(*
	Contract shared by span exporters. A processor offers a batch with export, which moves up to
	count of the oldest spans out of the processor's queue into the exporter without cloning
	them. The exporter owns the batch until free, which runs when the batch is delivered or
	failed, when the next batch is accepted, and when the exporter is destroyed.
	Concrete exporters advance delivery in tick and report through isBusy whether they can take
	another batch. Only ended spans reach an exporter.
*)
FUNCTION_BLOCK ABSTRACT FB_SpanExporter_Base
VAR
	_spans: FB_SpanQueue(maxCount:=0);
	_exportActive: BOOL;
	_callFailureReason: E_SpanExporterFailureReason;
END_VAR

(*
	Takes ownership of up to count of the oldest spans in spans. While busy it refuses with
	ACTIVE_EXPORT_IN_PROGRESS and leaves spans unchanged. A count of zero accepts nothing and
	succeeds.
*)
METHOD export : BOOL
VAR_IN_OUT
	spans: FB_SpanQueue;  // accepted spans are transferred out of this queue
END_VAR
VAR_INPUT
	count: UDINT;
END_VAR
VAR_OUTPUT
	failureReason: E_SpanExporterFailureReason;
END_VAR
VAR
	_queueFailureReason: E_SpanQueueFailureReason;
END_VAR
export := FALSE;
failureReason := E_SpanExporterFailureReason.NA;

IF THIS^.isBusy() THEN
	failureReason := E_SpanExporterFailureReason.ACTIVE_EXPORT_IN_PROGRESS;
	RETURN;
END_IF

// release a finished batch still held by the exporter before accepting the next one
THIS^.free();
IF NOT spans.transferTo(
	destination:=THIS^._spans,
	count:=count,
	failureReason=>_queueFailureReason
) THEN
	failureReason := E_SpanExporterFailureReason.QUEUE_TRANSFER_FAILURE;
	RETURN;
END_IF

THIS^._exportActive := THIS^._spans.count > 0;
export := TRUE;
END_METHOD

METHOD FB_Exit : BOOL
VAR_INPUT
	bInCopyCode: BOOL;
END_VAR
IF NOT bInCopyCode THEN
	THIS^.free();
END_IF
END_METHOD

(* Releases every span the exporter owns and clears the active export. *)
METHOD free
THIS^._spans.free();
THIS^._exportActive := FALSE;
END_METHOD

(* TRUE while the exporter cannot accept another batch. *)
METHOD ABSTRACT isBusy : BOOL
END_METHOD

(* Advances delivery of the accepted batch. Call it every scan. *)
METHOD ABSTRACT tick : BOOL
VAR_OUTPUT
	failureReason: E_SpanExporterFailureReason;
END_VAR
END_METHOD

END_FUNCTION_BLOCK

(* stored: Version 1.1.0.1
   POU FB_SpanExporter_Base: Id {7c2c489b-aca7-451b-ae42-a43cab088e9b}, SpecialFunc None
   Method export: Id {0626c578-cb2b-43ae-8054-5c85bcfdb916}
   Method FB_Exit: Id {e0fb3d50-e99d-4fc9-bacf-ab8571b068ba}
   Method free: Id {777bbfc3-1e9f-41b6-ba68-5ec6ed3a5b8c}
   Method isBusy: Id {becd6464-9b53-4e3d-8a80-79ff1418c346}
   Method tick: Id {67304bcf-08e8-4aac-bd2c-b5191c343fbc} *)
